// TIA Portal V21 export
DATA_BLOCK "TiaMcpComponentGate_1"   // DB2
VERSION : 0.1
// stored: AutoNumber false, DBAccessibleFromOPCUA true, DBAccessibleFromWebserver true, InstanceOfName TiaMcpComponentGate, InstanceOfType FB
"TiaMcpComponentGate"
   // VAR_INPUT
   //    Enable : Bool;
   // END_VAR
   // VAR_OUTPUT
   //    Active : Bool;
   // END_VAR
   // VAR
   //    State { S7_SetPoint := 'True'} : "TiaMcpComponentState";
   // END_VAR
BEGIN
END_DATA_BLOCK
